{attribute 'linkalways'}
{attribute 'no_explicit_call' := 'Use the methods of this class'}
{attribute 'enable_dynamic_creation'}
FUNCTION_BLOCK Accelerometer_Simulated IMPLEMENTS I_Accelerometer
VAR
	link : REFERENCE TO SimulatorLink;
END_VAR

METHOD FB_init : BOOL
VAR_INPUT
	bInitRetains : BOOL;
	bInCopyCode : BOOL;
	simulator : REFERENCE TO SimulatorLink;
END_VAR
link REF= simulator;
END_METHOD

PROPERTY AccelerationInMPerS2 : Vector3
GET
AccelerationInMPerS2 := SimulatorIo.feedback.accelerationInMPerS2;
END_GET
END_PROPERTY

PROPERTY TimestampInNs : ULINT
GET
TimestampInNs := SimulatorIo.feedback.timeInNs;
END_GET
END_PROPERTY

PROPERTY IsValid : BOOL
GET
IsValid := __ISVALIDREF(link) AND_THEN link.IsConnected;
END_GET
END_PROPERTY

END_FUNCTION_BLOCK

(* stored: Version 1.1.0.1, ProductVersion 3.1.4026.12
   POU Accelerometer_Simulated: Id {4c7be470-05ab-5175-8ee2-55f53b33fcd1}, SpecialFunc None
   Method FB_init: Id {8db6a0a0-9b3a-50be-af2c-5eaf94e8b1a3}
   Property AccelerationInMPerS2: Id {3cdf711d-364c-50fc-95bd-905692904ae6}
   Get Get: Id {4c3af306-ede9-5442-8072-437fdf85f2d3}
   Property TimestampInNs: Id {c7940b2a-d44f-5735-9ee7-c7cf5f4f8864}
   Get Get: Id {1105b718-f12c-5f89-a472-0749bd7c984b}
   Property IsValid: Id {dbbe89e6-0553-5096-8e51-77adf47f0320}
   Get Get: Id {42ce643a-0423-576e-bae9-c717efeaa091} *)
